Staubli VAL3: main.pgx

program main()
begin
  close(tCurrentTool)
  pPointRs.config.shoulder = lefty
  pPointRs2.config.shoulder = lefty
  mCurrentSpeed.tvel = 100.00
  mCurrentSpeed.blend = joint
  mCurrentSpeed.reach = 0.010
  mCurrentSpeed.leave = 0.010
  // Program TgtProg start
  // Program generated by RoboDK v6.0.7 for Staubli RX130B on XX/XX/XXXX 18:00:00
  // Using nominal kinematics.
  pPointRs.config.shoulder = righty
  call MoveLine(-607.850,543.849,363.215,136.262,30.757,-130.375)
  call MoveLine(-607.850,543.849,363.215,136.262,30.757,-130.375)
  pPointRs.config.shoulder = lefty
  call MoveLine(-607.850,543.849,363.215,136.262,30.757,-130.375)

  waitEndMove()
  // Program TgtProg end

end
